Fanuc KAREL source: KT00204.KL

PROGRAM KT00204
%NOLOCKGROUP
VAR
  I1: INTEGER
  I2: INTEGER
  OUT: INTEGER
BEGIN
  I1 = 2
  I2 = 3
  I1 = 2
  I2 = 3
  OUT = I1 AND I2
END KT00204
